FUNCTION_BLOCK PUBLIC TcoRtc IMPLEMENTS ITcoRtc
VAR
	{attribute 'hide'}
	_isValid							:	BOOL := FALSE;
	{attribute 'hide'}
	_state								:	UINT;
	{attribute 'hide'}
	_TimeZoneID							:	Tc2_EtherCAT.Tc2_Utilities.E_TimeZoneID;
	{attribute 'hide'}
	_NT_GetLocalTime					: 	Tc2_EtherCAT.Tc2_Utilities.NT_GetTime;
	{attribute 'hide'}
	_FB_TzSpecificLocalTimeToSystemTime :	Tc2_EtherCAT.Tc2_Utilities.FB_TzSpecificLocalTimeToSystemTime;
	{attribute 'hide'}
	_RTC_EX2							:	Tc2_EtherCAT.Tc2_Utilities.RTC_EX2;
	{attribute 'hide'}
	_PDT	 							:	Tc2_EtherCAT.Tc2_Utilities.TIMESTRUCT;	
	{attribute 'hide'}
	_LocalTime 							:	Tc2_EtherCAT.Tc2_Utilities.TIMESTRUCT;
	{attribute clr [ReadOnly()]}
	_LocalTimeDT						:	DATE_AND_TIME;
	{attribute 'hide'}
	_UTCTime 							:	Tc2_EtherCAT.Tc2_Utilities.TIMESTRUCT;
	{attribute clr [ReadOnly()]}
	_UTCTimeDT							:	DATE_AND_TIME;
END_VAR

PROPERTY IsSynchronized : BOOL
GET
IsSynchronized :=  RtcPrg._isSynchronized;
END_GET
END_PROPERTY

PROPERTY IsValid : BOOL
GET
IsValid := _isValid;
END_GET
END_PROPERTY

METHOD NowLocal : DATE_AND_TIME
IF _isValid THEN
	NowLocal := _LocalTimeDT;
END_IF
END_METHOD

METHOD NowLocalAsTIMESTRUCT : Tc2_EtherCAT.Tc2_Utilities.TIMESTRUCT
IF _isValid THEN
	NowLocalAsTIMESTRUCT := _LocalTime;
END_IF
END_METHOD

METHOD NowUTC : DATE_AND_TIME
IF _isValid THEN
	NowUTC := _UTCTimeDT;
END_IF
END_METHOD

METHOD NowUTCAsTIMESTRUCT : Tc2_EtherCAT.Tc2_Utilities.TIMESTRUCT
IF _isValid THEN
	NowUTCAsTIMESTRUCT := _UTCTime;
END_IF
END_METHOD

METHOD TickClock : ULINT
TickClock := Tc2_EtherCAT.F_GetActualDcTime64();
END_METHOD

METHOD PROTECTED Update
VAR
	_diffToLastSyncInSeconds : LINT;
END_VAR
IF _state = 0 THEN
//	_isValid := FALSE;
	_NT_GetLocalTime(NETID := '127.0.0.1.1.1', START := TRUE);
	IF _NT_GetLocalTime.BUSY AND NOT _NT_GetLocalTime.ERR THEN 
		_state := _state + 10;
	END_IF
END_IF
	
IF _state = 10 THEN
	_NT_GetLocalTime(START := FALSE);
	IF NOT _NT_GetLocalTime.BUSY AND NOT _NT_GetLocalTime.ERR THEN 
		_state := _state + 10;
	END_IF
END_IF

IF _state = 20 THEN
	_NT_GetLocalTime(START := FALSE);
		
	_PDT := _NT_GetLocalTime.TIMESTR;

	_isValid := TRUE;
END_IF

_RTC_EX2(EN := _isValid, PDT := _PDT);

_diffToLastSyncInSeconds := ABS(ULINT_TO_LINT(Tc2_EtherCAT.SYSTEMTIME_TO_DCTIME64(_RTC_EX2.CDT,0,0) - Tc2_EtherCAT.SYSTEMTIME_TO_DCTIME64(RtcPrg._LastSyncTimeStampInLocalTime,0,0)))/1000000000;

IF _state >= 20 AND RtcPrg._RtcSynchParams.doSynch AND _diffToLastSyncInSeconds >=RtcPrg._RtcSynchParams.syncPeriod THEN
	_state := 0;
END_IF

_LocalTime := _RTC_EX2.CDT;
_LocalTimeDT := Tc2_EtherCAT.Tc2_Utilities.SYSTEMTIME_TO_DT(_LocalTime);

IF RtcPrg._isSynchronized THEN
	_FB_TzSpecificLocalTimeToSystemTime(in 		:=	_LocalTime,
										tzInfo 	:=	RtcPrg._TimeZoneInformation,
										out		=>	_UTCTime,
										eTzID	=>	_TimeZoneID);
	_UTCTimeDT := Tc2_EtherCAT.Tc2_Utilities.SYSTEMTIME_TO_DT(_UTCTime);
END_IF
END_METHOD

METHOD INTERNAL UpdateInternal
THIS^.Update();
END_METHOD

END_FUNCTION_BLOCK

(* stored: Version 1.1.0.1
   POU TcoRtc: Id {44984f17-252b-05a5-3965-3576c168912a}, SpecialFunc None
   Property IsSynchronized: Id {281d422f-3fd6-08a1-39a9-839854b5b3de}
   Get Get: Id {56a732cd-dbfe-0b14-1254-ee3c7eed7852}
   Property IsValid: Id {0b73d0fb-6a2d-0c9e-3da7-384d62e156b5}
   Get Get: Id {f1495f6e-f4ab-08bd-138d-164d6df2166a}
   Method NowLocal: Id {ba634665-0212-047c-1c1d-6ebb5a5f30b5}
   Method NowLocalAsTIMESTRUCT: Id {e9fe0ffa-a159-017e-3bd5-9e67f37e7fa9}
   Method NowUTC: Id {34a4b82c-d3a2-0332-3148-6e27e32eec88}
   Method NowUTCAsTIMESTRUCT: Id {6c922f94-0952-07e6-0cac-83326b01c28c}
   Method TickClock: Id {1cdfb043-4f81-0904-37ac-2a0334c75a58}
   Method Update: Id {0bf459e2-db45-0e5b-3d87-31081b5a02e2}
   Method UpdateInternal: Id {c570233f-a171-005d-1421-aec37fed972f} *)
